// TIA Portal V20 export
// export: Created 2000-01-01T00:00:00.0000000Z, ExportSetting None
FUNCTION "FC_Rung" : Void   // FC42, LAD
{ S7_Optimized_Access := 'TRUE' }
   VAR_INPUT
      Local : Int;
   END_VAR
   VAR_TEMP   // added for the SCL form of the ladder/FBD networks
      _w1 : Bool;
   END_VAR
BEGIN

REGION Network 1
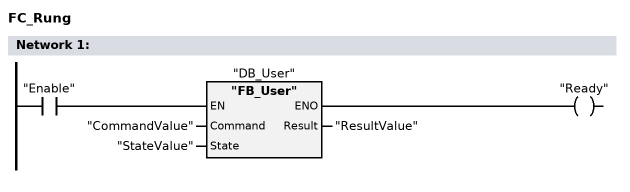
   RUNG wire#powerrail
      Contact( "Enable" )
      "DB_User"(Command := "CommandValue", State := "StateValue", Result => "ResultValue")
      Coil( "Ready" )
   END_RUNG
   // the same network as SCL:
   "DB_User"(EN := "Enable",   // "FB_User"
             Command := "CommandValue",
             State := "StateValue",
             Result => "ResultValue",
             ENO => #_w1);
   "Ready" := #_w1;
END_REGION
END_FUNCTION
